Fanuc KAREL source: KA00164.KL

PROGRAM KA00164
%NOLOCKGROUP
VAR
  SRC: ARRAY[4] OF BOOLEAN
  DST: ARRAY[4] OF REAL
BEGIN
  DST = SRC
END KA00164
